Fanuc KAREL source: kt00304.KL

PROGRAM KT00304
%STACKSIZE=65535
%PRIORITY=65535
%NOLOCKGROUP
VAR
Y1 : ARRAY[2] OF BYTE
R2 : REAL
OUT : BOOLEAN
BEGIN
Y1[1]=2
R2=3.0
OUT=(R2 <> (Y1[1]))
END KT00304
